FUNCTION_BLOCK FB_Tc
VAR_INPUT
    bEnable : BOOL;
END_VAR
VAR
    nValue : INT;
    nForgotten : INT; // PLCA-Q001
END_VAR

IF bEnable THEN
    nValue := nValue + 1;
END_IF

END_FUNCTION_BLOCK

(* stored: Version 1.1.0.1, ProductVersion 3.1.4024.12
   POU FB_Tc: Id {11111111-2222-3333-4444-555555555555}, SpecialFunc None *)
